Fanuc KAREL source: ka00225.KL

PROGRAM KA00225
%STACKSIZE=65535
%PRIORITY=65535
%NOLOCKGROUP
VAR
SRC : ARRAY[4] OF JOINTPOS9
DST : ARRAY[4] OF JOINTPOS9
BEGIN
-- UNRESOLVED_PC line 7 opcodes [22 22 1E] marker_code=0
END KA00225
